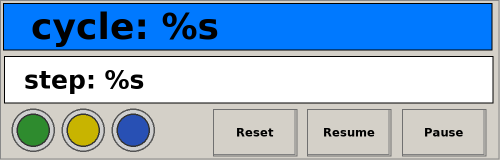
VISUALIZATION vis_Cycle_Control  // 500x160
VAR_IN_OUT
	fb: FB_SFC_Cycle;
END_VAR
VAR_INPUT
	sName: STRING:='Cycle name';
END_VAR
    Lamp1 (8,105 50x50), tooltip "Ready", variable: fb.bReady, style: Lamp-Lamp1-Green
    Lamp1 (108,105 50x50), tooltip "Done", variable: fb.bDone, style: Lamp-Lamp1-Blue
    Lamp1 (58,105 50x50), tooltip "Run", variable: fb.bRun, style: Lamp-Lamp1-Yellow
    RoundedRectangle (3,3 489x47), "cycle: %s", tooltip "POU name: %s", text variable: sName
        p4168582468: fb.refSFC.SFCErrorPOU
    RoundedRectangle (4,56 489x47), "step: %s", text variable: fb.refSFC.SFCCurrentStep, colour toggle: fb.ErrorSFC
    Button (213,109 84x47), "Reset"
        tap fb.bInit
    Button (307,109 84x47), "Resume", colour toggle: fb.ErrorSFC
        toggle fb.refSFC.SFCQuitError
    Button (402,109 84x47), "Pause", colour toggle: fb.refSFC.SFCPause
        toggle fb.refSFC.SFCPause
END_VISUALIZATION

(* stored: Version 1.1.0.1, ProductVersion 3.1.4024.12
   Visu vis_Cycle_Control: Id {fd349829-2291-4f50-a259-aa5f8002aba7} *)
